FUNCTION FC 1 : VOID
NETWORK
      A I 0.0
END_FUNCTION
